// TIA Portal V20 export
// export: Created 2026-10-19T18:45:17.0120055Z, ExportSetting None, DisplayName Totally Integrated Automation Portal, DisplayVersion V20 Update 6, DisplayName TIA Portal Openness, DisplayVersion V20 Update 6, DisplayName TIA Portal Version Control Interface, DisplayVersion V20 Update 6, DisplayName SINAMICS Startdrive Advanced, DisplayVersion V20 SP1, DisplayName SINAMICS Startdrive G130, G150, S120, S150, SINAMICS MV, G220, S200, S210, DisplayVersion V20 SP1, DisplayName SINAMICS Startdrive G110M, G120, G120C, G120D, G120P, G115D, DisplayVersion V20 SP1, DisplayName STEP 7 Professional, DisplayVersion V20 Update 6, DisplayName STEP 7 Safety, DisplayVersion V20 Update 2, DisplayName WinCC Basic/Comfort/Advanced, DisplayVersion V20 Update 6, DisplayName WinCC Unified, DisplayVersion V20 Update 6
VAR_GLOBAL   // PLC tag table "PopUp_Screens"
   LE_Speed AT %MW710 : Int;
   LE_Warnings AT %MW714 : Int;
   LE_Status AT %MW702 : UInt;
   LE_Quality_Value AT %MB716 : Byte;
   LE_X_Unsafe_Position AT %MD706 : DInt;
   LE_Quality_Decoded_Codes AT %MB724 : Byte;
   LE_Bypass AT %M704.0 : Bool;
   AE_Speed AT %MW96 : Int;
   AE_Status_2 AT %MW100 : UInt;
   AE_Control_Word_2 AT %MW86 : UInt;
   AE_Position_1 AT %MD88 : DInt;
   AE_Position_2 AT %MD92 : DInt;
   AE_Status_1 AT %MW98 : UInt;
   AE_Control_Word_1 AT %MW156 : UInt;
   BCD_Disable_Trigger_HMI AT %M1156.2 : Bool;
   BCD_Enable_Trigger_HMI AT %M1156.1 : Bool;
   BCD_Error_HMI AT %M1156.3 : Bool;
   BCD_Start_Comm_Test_HMI AT %M1156.0 : Bool;
   BCD_Test_Ok_HMI AT %M1156.4 : Bool;
   BCD_Execute_Function AT %M1156.5 : Bool;
   BCD_RdDone AT %M1156.7 : Bool;
   BCD_ReqDone AT %M1157.0 : Bool;
   BCD_ReqBusy AT %M1157.1 : Bool;
END_VAR
